Fanuc KAREL source: kt00168.KL

-- PROVISIONAL review KL for V940-1; original PC SHA256 4713e584fb60d987ab15db2235d690936828284fc9913c6a319b1796be5a2440
-- Incomplete behavior may be omitted. Consult companion uncertainty JSON. Do not deploy.
PROGRAM KT00168
%NOLOCKGROUP
VAR
  I1 : INTEGER
  OUT : REAL
-- UNRESOLVED_DECL H2 type=002017
BEGIN
  -- V9_ZERO_TABLE_METADATA_HINT layout=0001; no indexed target words; source/name/runtime held
  -- UNRESOLVED_PC offsets 5-16; opcodes 2E,23
  -- UNRESOLVED_PC offsets 21-35; opcodes 2E,22,9D,33,B4
  -- UNRESOLVED_PC offsets 40-63; opcodes 21,22,9D,33,B3,56,64,23
  -- UNRESOLVED_PC offsets 68-72; opcodes 7F
END KT00168
